FUNCTION_BLOCK FB_RMP_W
VAR_INPUT
	bEnable			:BOOL := TRUE;	(* Enable input *)
	bDirection		:BOOL := TRUE;	(* Direction Up = TRUE, means up *)
	bSet 			:BOOL;			(* Set input *)
	bReset 			:BOOL;			(* Reset input *)
	tRampTime	 	:TIME;			(* Duration of a ramp 0..65535 *)
END_VAR
VAR_OUTPUT
	wRVOut 			:WORD;			(* Ramp output *)
	bBusy 			:BOOL;			(* TRUE, when ramp is running *)
	bLowLevel 		:BOOL;			(* Minimum output value is reached *)
	bHighLevel 		:BOOL;			(* Maximum output value is reached *)
END_VAR
VAR
	fbRamp 			: _RMP_W;
END_VAR

(*
version 2.0	23. oct. 2008
programmer 	oscat
tested BY	oscat

this ramp generator generates a Word wide ramp with 65535 steps
the generator has an asynchronous set and reset
the ramp is controlled by PT which is the total ramp time for a full sweep from 0..65535
an UD input controlls the direction Up or Down and the E input enables the ramp generation
a busy output indicates that the ramp is running, busy false means output is stable.
the outputs low and high will be true when the output has reached its max or min value.

RMP_W is a ramp generator with 16-bit (2 bytes) resolution. The ramp of
0.. 65535 is divided into a maximum of 65536 steps and run in a time of
PT once complete. An enable signal E switches the ramp generator on or
of. An asynchronous reset sets each time the output to 0, and a pulse at
the Set input sets the output to 65535. With the UD input, the direction UP
(UD = TRUE) or DOWN (UD = FALSE) is defined. The output of BUSY =
TRUE indicates that a ramp is active. BUSY = FALSE means the output is
stable. The outputs HIGH and LOW gets TRUE, the output OUT reaches the
lower or upper limit (0 and 65535).
At setting of PT is to be noted that a PLC with 5 ms cycle time needs
65536*5 = 327 seconds for a ramp. If the PT is the time defined shorter
than the cycle time 65536, the edge is translated in correspondingly larger
steps. The ramp is constructed in this case with less than 256 steps
per cycle. PT may be T#0s, then the output switched between minimum
and maximum value back and forth.
For a detailed description, see the module RMP_B. The function is absolutely
identical except that the output OUT 8-bit wide instead of 16 bit.
*)

(* Generate ramp *)
fbRamp(
	bEnable := bEnable,
	bDirection := bDirection,
	tFullRmpTime := tRampTime,
	wRamp := wRVOut
);

(* Set or Reset operation *)
IF bReset
THEN
	wRVOut := 0;
ELSIF bSet
THEN
	wRVOut := 65535;
END_IF;

(* Checks for outputs stable and reset or set busy flag *)
bLowLevel := wRVOut = 0;
bHighLevel := wRVOut = 65535;
bBusy := bEnable
	        AND NOT (bLowLevel OR bHighLevel);

END_FUNCTION_BLOCK

(* stored: Version 1.1.0.1, ProductVersion 3.1.4024.15
   POU FB_RMP_W: Id {9761fe48-60a2-44d2-aa18-06ef6f412b67}, SpecialFunc None *)
